Staubli VAL3: getFrameID.pgx

public program getFrameID(string x_sKey, num& x_nFrameID)
begin
  x_nFrameID=trajTemp:tTrajItem[x_sKey].nFrameIndex
end
